// Mitsubishi GX Works2 project: 261012_저속+고속타이머   PLC: Q03UDV

PROGRAM MAIN
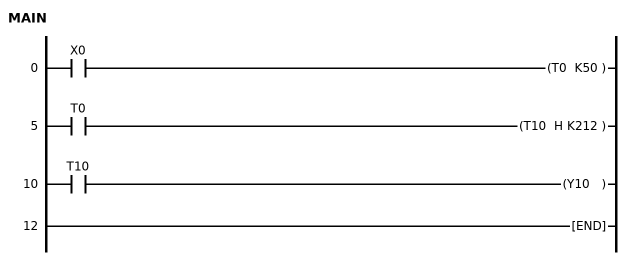
0     LD      X0
      OUT     T0 K50
5     LD      T0
      OUTH    T10 K212
10    LD      T10
      OUT     Y10
12    END
END_PROGRAM
